// TIA Portal V19 export
DATA_BLOCK "Sim_SMOutputs_DB"   // DB9
// stored: InstanceOfName Sim_SMOutputs, InstanceOfType FB
"Sim_SMOutputs"
   // VAR
   //    VaccumPID { ExternalAccessible := 'False'; ExternalVisible := 'False'; ExternalWritable := 'False'} : "PidL";
   //    SteamPID { S7_SetPoint := 'True'} : "PidL";
   //    SimularDelay { S7_SetPoint := 'True'} : TON_TIME;
   //    FeedPID { S7_SetPoint := 'True'} : "PidL";
   //    LiSet : Bool := FALSE;
   //    LiSetM : Bool := FALSE;
   //    LevelInit : Real := 0.0;
   //    BrixInit : Real := 0.0;
   // END_VAR
BEGIN
   VaccumPID.AutModLi := TRUE;
   VaccumPID.ManModLi := FALSE;
   VaccumPID.LocModLi := FALSE;
   VaccumPID.OosModLi := FALSE;
   VaccumPID.ModLiOp := TRUE;
   VaccumPID.ResetLi := FALSE;
   VaccumPID.SPModLiOp := FALSE;
   VaccumPID.ExtModLi := FALSE;
   VaccumPID.IntModLi := FALSE;
   VaccumPID.PV := 950.0145;
   VaccumPID.PV_Norm.High := 2000.0;
   VaccumPID.PV_Norm.Low := 0.0;
   VaccumPID.MV_Norm.High := 100.0;
   VaccumPID.MV_Norm.Low := 0.0;
   VaccumPID.PV_Scale.High := 2000.0;
   VaccumPID.PV_Scale.Low := 0.0;
   VaccumPID.SPExt := 0.0;
   VaccumPID.SP_HiLim := 1000.0;
   VaccumPID.SP_LoLim := 0.0;
   VaccumPID.MV_HiLim := 100.0;
   VaccumPID.MV_LoLim := 0.0;
   VaccumPID.OosSafeMV := 0.0;
   VaccumPID.PV_unit := 1342;
   VaccumPID.MV_unit := 1342;
   VaccumPID.DataHMI.identName := '';
   VaccumPID.DataHMI.comment := '';
   VaccumPID.DataHMI.AutModOp := TRUE;
   VaccumPID.DataHMI.ManModOp := FALSE;
   VaccumPID.DataHMI.LocModOp := FALSE;
   VaccumPID.DataHMI.OosModOp := FALSE;
   VaccumPID.DataHMI.ResetOp := FALSE;
   VaccumPID.DataHMI.MonitorOn := FALSE;
   VaccumPID.DataHMI.ExtModOp := FALSE;
   VaccumPID.DataHMI.IntModOp := FALSE;
   VaccumPID.DataHMI.SpInt := 100.0;
   VaccumPID.DataHMI.Man := 0.0;
   VaccumPID.DataHMI.PermissionLog.AutModOpEn := FALSE;
   VaccumPID.DataHMI.PermissionLog.ManModOpEn := FALSE;
   VaccumPID.DataHMI.PermissionLog.LocModOpEn := FALSE;
   VaccumPID.DataHMI.PermissionLog.OosModOpEn := FALSE;
   VaccumPID.DataHMI.PermissionLog.ResetOpEn := TRUE;
   VaccumPID.DataHMI.PermissionLog.ExtModOpEn := FALSE;
   VaccumPID.DataHMI.PermissionLog.IntModOpEn := FALSE;
   VaccumPID.DataHMI.PermissionLog.Alarms.MsgSupEn := FALSE;
   VaccumPID.DataHMI.PermissionLog.Alarms.HiAlmSupEn := FALSE;
   VaccumPID.DataHMI.PermissionLog.Alarms.HiWrnSupEn := FALSE;
   VaccumPID.DataHMI.PermissionLog.Alarms.LoWrnSupEn := FALSE;
   VaccumPID.DataHMI.PermissionLog.Alarms.LoAlmSupEn := FALSE;
   VaccumPID.DataHMI.Status.OosAct := FALSE;
   VaccumPID.DataHMI.Status.LocAct := FALSE;
   VaccumPID.DataHMI.Status.ManAct := FALSE;
   VaccumPID.DataHMI.Status.AutAct := TRUE;
   VaccumPID.DataHMI.Status.SpExtAct := FALSE;
   VaccumPID.DataHMI.Status.Protection := FALSE;
   VaccumPID.DataHMI.Status.Intlock := TRUE;
   VaccumPID.DataHMI.Status.Permit := TRUE;
   VaccumPID.DataHMI.Status.TrackAct := TRUE;
   VaccumPID.DataHMI.Status.SP := 100.0;
   VaccumPID.DataHMI.Status.PV := 950.0145;
   VaccumPID.DataHMI.Status.ER := -845.0145;
   VaccumPID.DataHMI.Status.MV := 0.0;
   VaccumPID.DataHMI.Status.PVOpScale.High := 2000.0;
   VaccumPID.DataHMI.Status.PVOpScale.Low := 0.0;
   VaccumPID.DataHMI.Status.MVOpScale.High := 100.0;
   VaccumPID.DataHMI.Status.MVOpScale.Low := 0.0;
   VaccumPID.DataHMI.Status.SPIntLim.High := 0.0;
   VaccumPID.DataHMI.Status.SPIntLim.Low := 0.0;
   VaccumPID.DataHMI.Status.PV_unit := 1342;
   VaccumPID.DataHMI.Status.MV_unit := 1342;
   VaccumPID.DataHMI.PIDConfig.NegGain := TRUE;
   VaccumPID.DataHMI.PIDConfig.P_Sel := TRUE;
   VaccumPID.DataHMI.PIDConfig.I_Sel := TRUE;
   VaccumPID.DataHMI.PIDConfig.D_Sel := FALSE;
   VaccumPID.DataHMI.PIDConfig.Gain := -2.0;
   VaccumPID.DataHMI.PIDConfig.Ti := 80.0;
   VaccumPID.DataHMI.PIDConfig.Td := 0.0;
   VaccumPID.DataHMI.PIDConfig.DeadBW := 5.0;
   VaccumPID.DataHMI.Alarms.identName := '';
   VaccumPID.DataHMI.Alarms.comment := '';
   VaccumPID.DataHMI.Alarms.MsgSupOp := FALSE;
   VaccumPID.DataHMI.Alarms.PVScale.High := 2000.0;
   VaccumPID.DataHMI.Alarms.PVScale.Low := 0.0;
   VaccumPID.DataHMI.Alarms.HiAlmSupOp := FALSE;
   VaccumPID.DataHMI.Alarms.HiWrnSupOp := FALSE;
   VaccumPID.DataHMI.Alarms.LoWrnSupOp := FALSE;
   VaccumPID.DataHMI.Alarms.LoAlmSupOp := FALSE;
   VaccumPID.DataHMI.Alarms.PermissionLog.MsgSupEn := FALSE;
   VaccumPID.DataHMI.Alarms.PermissionLog.HiAlmSupEn := TRUE;
   VaccumPID.DataHMI.Alarms.PermissionLog.HiWrnSupEn := TRUE;
   VaccumPID.DataHMI.Alarms.PermissionLog.LoWrnSupEn := TRUE;
   VaccumPID.DataHMI.Alarms.PermissionLog.LoAlmSupEn := TRUE;
   VaccumPID.DataHMI.Alarms.Status.PV := 950.0145;
   VaccumPID.DataHMI.Alarms.Status.PV_unit := 1342;
   VaccumPID.DataHMI.Alarms.Status.PV_HiAlm := TRUE;
   VaccumPID.DataHMI.Alarms.Status.PV_HiWrn := TRUE;
   VaccumPID.DataHMI.Alarms.Status.PV_LoWrn := FALSE;
   VaccumPID.DataHMI.Alarms.Status.PV_LoAlm := FALSE;
   VaccumPID.DataHMI.Alarms.Status.MsgSup := FALSE;
   VaccumPID.Feature.Startup := TRUE;
   VaccumPID.Feature.MSSOff := TRUE;
   VaccumPID.Feature.FltOff := TRUE;
   VaccumPID.Feature.LocalMod := FALSE;
   VaccumPID.Permission.AutModOpEn := TRUE;
   VaccumPID.Permission.ManModOpEn := TRUE;
   VaccumPID.Permission.LocModOpEn := FALSE;
   VaccumPID.Permission.OosModOpEn := FALSE;
   VaccumPID.Permission.ResetOpEn := TRUE;
   VaccumPID.Permission.ExtModOpEn := FALSE;
   VaccumPID.Permission.IntModOpEn := TRUE;
   VaccumPID.Permission.Alarms.MsgSupEn := TRUE;
   VaccumPID.Permission.Alarms.HiAlmSupEn := TRUE;
   VaccumPID.Permission.Alarms.HiWrnSupEn := TRUE;
   VaccumPID.Permission.Alarms.LoWrnSupEn := TRUE;
   VaccumPID.Permission.Alarms.LoAlmSupEn := TRUE;
   VaccumPID.MSS := TRUE;
   VaccumPID.Trip := FALSE;
   VaccumPID.Permit := TRUE;
   VaccumPID.Intlock := TRUE;
   VaccumPID.Protect := TRUE;
   VaccumPID.TrackOn := TRUE;
   VaccumPID.Rbk := 0.0;
   VaccumPID.RbkHiTol := 3.0;
   VaccumPID.RbkLoTol := 3.0;
   VaccumPID.RbkMonTime := T#3S;
   VaccumPID.TrackVal := 0.0;
   VaccumPID.RunUpCyc := 3;
   VaccumPID.DisV := 0.0;
   VaccumPID.HiAlm := 95.0;
   VaccumPID.HiWrn := 90.0;
   VaccumPID.LoWrn := 10.0;
   VaccumPID.LoAlm := 5.0;
   VaccumPID.Hyst := 5.0;
   VaccumPID.AutAct := TRUE;
   VaccumPID.ManAct := FALSE;
   VaccumPID.LocAct := FALSE;
   VaccumPID.OosAct := FALSE;
   VaccumPID.MsgSup := TRUE;
   VaccumPID.AlarmError := FALSE;
   VaccumPID.MV := 0.0;
   VaccumPID.SPExtAct := FALSE;
   VaccumPID.SP := 100.0;
   VaccumPID.ER := -845.0145;
   VaccumPID.PVH_Alm := TRUE;
   VaccumPID.PVH_Wrn := TRUE;
   VaccumPID.PVL_Wrn := FALSE;
   VaccumPID.PVL_Alm := FALSE;
   VaccumPID.controller.COM_RST := FALSE;
   VaccumPID.controller.MAN_ON := TRUE;
   VaccumPID.controller.PVPER_ON := FALSE;
   VaccumPID.controller.P_SEL := TRUE;
   VaccumPID.controller.I_SEL := TRUE;
   VaccumPID.controller.INT_HOLD := FALSE;
   VaccumPID.controller.I_ITL_ON := FALSE;
   VaccumPID.controller.D_SEL := FALSE;
   VaccumPID.controller.CYCLE := T#200MS;
   VaccumPID.controller.SP_INT := 5.0;
   VaccumPID.controller.PV_IN := 47.50072;
   VaccumPID.controller.PV_PER := 16#0000;
   VaccumPID.controller.MAN := 0.0;
   VaccumPID.controller.GAIN := -2.0;
   VaccumPID.controller.TI := T#1M_20S;
   VaccumPID.controller.TD := T#10S;
   VaccumPID.controller.TM_LAG := T#2S;
   VaccumPID.controller.DEADB_W := 0.25;
   VaccumPID.controller.LMN_HLM := 100.0;
   VaccumPID.controller.LMN_LLM := 0.0;
   VaccumPID.controller.PV_FAC := 1.0;
   VaccumPID.controller.PV_OFF := 0.0;
   VaccumPID.controller.LMN_FAC := 1.0;
   VaccumPID.controller.LMN_OFF := 0.0;
   VaccumPID.controller.I_ITLVAL := 0.0;
   VaccumPID.controller.DISV := 0.0;
   VaccumPID.controller.LMN := 0.0;
   VaccumPID.controller.LMN_PER := 16#0000;
   VaccumPID.controller.QLMN_HLM := FALSE;
   VaccumPID.controller.QLMN_LLM := TRUE;
   VaccumPID.controller.LMN_P := 84.50145;
   VaccumPID.controller.LMN_I := -84.50145;
   VaccumPID.controller.LMN_D := 0.0;
   VaccumPID.controller.PV := 47.50072;
   VaccumPID.controller.ER := -42.25072;
   VaccumPID.controller.sInvAlt := 84.50145;
   VaccumPID.controller.sIanteilAlt := -84.50145;
   VaccumPID.controller.sRestInt := 0.0;
   VaccumPID.controller.sRestDif := 0.0;
   VaccumPID.controller.sRueck := 84.50145;
   VaccumPID.controller.sLmn := 0.0;
   VaccumPID.controller.sbArwHLmOn := FALSE;
   VaccumPID.controller.sbArwLLmOn := TRUE;
   VaccumPID.controller.sbILimOn := TRUE;
   VaccumPID.ModSelInt := 2;
   VaccumPID.stRestart := FALSE;
   VaccumPID.ResetLiLogic := FALSE;
   VaccumPID.ResetResult := FALSE;
   VaccumPID.stResetLiLogic := FALSE;
   VaccumPID.stMonErr := FALSE;
   VaccumPID.stTripErr := FALSE;
   VaccumPID.stProtErr := FALSE;
   VaccumPID.stMSS := FALSE;
   VaccumPID.stProt := FALSE;
   VaccumPID.stTrip := FALSE;
   VaccumPID.stLockFault := FALSE;
   VaccumPID.stRun := FALSE;
   VaccumPID.stExtMod := FALSE;
   VaccumPID.stAutoLogic := FALSE;
   VaccumPID.RuntimeMem := 16#0000_07DF_2C3D_9711;
   VaccumPID.RuntimeS := 0.200026255103497;
   VaccumPID.PVMon.Feature.Startup := TRUE;
   VaccumPID.PVMon.Enable := TRUE;
   VaccumPID.PVMon.Permission.MsgSupEn := TRUE;
   VaccumPID.PVMon.Permission.HiAlmSupEn := TRUE;
   VaccumPID.PVMon.Permission.HiWrnSupEn := TRUE;
   VaccumPID.PVMon.Permission.LoWrnSupEn := TRUE;
   VaccumPID.PVMon.Permission.LoAlmSupEn := TRUE;
   VaccumPID.PVMon.DataHMI.identName := '';
   VaccumPID.PVMon.DataHMI.comment := '';
   VaccumPID.PVMon.DataHMI.MsgSupOp := FALSE;
   VaccumPID.PVMon.DataHMI.PVScale.High := 2000.0;
   VaccumPID.PVMon.DataHMI.PVScale.Low := 0.0;
   VaccumPID.PVMon.DataHMI.HiAlmSupOp := FALSE;
   VaccumPID.PVMon.DataHMI.HiWrnSupOp := FALSE;
   VaccumPID.PVMon.DataHMI.LoWrnSupOp := FALSE;
   VaccumPID.PVMon.DataHMI.LoAlmSupOp := FALSE;
   VaccumPID.PVMon.DataHMI.PermissionLog.MsgSupEn := FALSE;
   VaccumPID.PVMon.DataHMI.PermissionLog.HiAlmSupEn := TRUE;
   VaccumPID.PVMon.DataHMI.PermissionLog.HiWrnSupEn := TRUE;
   VaccumPID.PVMon.DataHMI.PermissionLog.LoWrnSupEn := TRUE;
   VaccumPID.PVMon.DataHMI.PermissionLog.LoAlmSupEn := TRUE;
   VaccumPID.PVMon.DataHMI.Status.PV := 950.0145;
   VaccumPID.PVMon.DataHMI.Status.PV_unit := 1342;
   VaccumPID.PVMon.DataHMI.Status.PV_HiAlm := TRUE;
   VaccumPID.PVMon.DataHMI.Status.PV_HiWrn := TRUE;
   VaccumPID.PVMon.DataHMI.Status.PV_LoWrn := FALSE;
   VaccumPID.PVMon.DataHMI.Status.PV_LoAlm := FALSE;
   VaccumPID.PVMon.DataHMI.Status.MsgSup := FALSE;
   VaccumPID.PVMon.RunUpCyc := 3;
   VaccumPID.PVMon.PV := 950.0145;
   VaccumPID.PVMon.HiAlm := 95.0;
   VaccumPID.PVMon.HiWrn := 90.0;
   VaccumPID.PVMon.LoWrn := 10.0;
   VaccumPID.PVMon.LoAlm := 5.0;
   VaccumPID.PVMon.Hyst := 5.0;
   VaccumPID.PVMon.PV_unit := 1342;
   VaccumPID.PVMon.MsgErr := FALSE;
   VaccumPID.PVMon.MsgSup := FALSE;
   VaccumPID.PVMon.PVH_Alm := TRUE;
   VaccumPID.PVMon.PVH_Wrn := TRUE;
   VaccumPID.PVMon.PVL_Wrn := FALSE;
   VaccumPID.PVMon.PVL_Alm := FALSE;
   VaccumPID.PVMon.stRestart := FALSE;
   VaccumPID.PVMon.RunUpCounter := 0;
   VaccumPID.PVMon.pSIG1 := TRUE;
   VaccumPID.PVMon.pSIG2 := TRUE;
   VaccumPID.PVMon.pSIG3 := FALSE;
   VaccumPID.PVMon.pSIG4 := FALSE;
   VaccumPID.PVMon.pAlarm := TRUE;
   VaccumPID.RunUpCounter := 0;
   VaccumPID.pAlarm := TRUE;
   VaccumPID.stMSSErr := FALSE;
   VaccumPID.SPMod := FALSE;
   VaccumPID.SPSelInt := 0;
   VaccumPID.stErr := FALSE;
   VaccumPID.stDivErr := FALSE;
   VaccumPID.stNegGain := TRUE;
   VaccumPID.stGain := -2.0;
   VaccumPID.stTi := 0.0;
   VaccumPID.stTd := 0.0;
   VaccumPID.stPIDConfig.NegGain := TRUE;
   VaccumPID.stPIDConfig.P_Sel := TRUE;
   VaccumPID.stPIDConfig.I_Sel := TRUE;
   VaccumPID.stPIDConfig.D_Sel := FALSE;
   VaccumPID.stPIDConfig.Gain := -2.0;
   VaccumPID.stPIDConfig.Ti := 80.0;
   VaccumPID.stPIDConfig.Td := 0.0;
   VaccumPID.stPIDConfig.DeadBW := 5.0;
   VaccumPID.RbkMonitorTimer.PT := T#0MS;
   VaccumPID.RbkMonitorTimer.IN := FALSE;
   SteamPID.AutModLi := TRUE;
   SteamPID.ManModLi := FALSE;
   SteamPID.LocModLi := FALSE;
   SteamPID.OosModLi := FALSE;
   SteamPID.ModLiOp := TRUE;
   SteamPID.ResetLi := FALSE;
   SteamPID.SPModLiOp := TRUE;
   SteamPID.ExtModLi := TRUE;
   SteamPID.IntModLi := FALSE;
   SteamPID.PV := 0.0;
   SteamPID.PV_Norm.High := 100.0;
   SteamPID.PV_Norm.Low := 0.0;
   SteamPID.MV_Norm.High := 100.0;
   SteamPID.MV_Norm.Low := 0.0;
   SteamPID.PV_Scale.High := 100.0;
   SteamPID.PV_Scale.Low := 0.0;
   SteamPID.SPExt := 80.0;
   SteamPID.SP_HiLim := 100.0;
   SteamPID.SP_LoLim := 0.0;
   SteamPID.MV_HiLim := 100.0;
   SteamPID.MV_LoLim := 0.0;
   SteamPID.OosSafeMV := 0.0;
   SteamPID.PV_unit := 1342;
   SteamPID.MV_unit := 1342;
   SteamPID.DataHMI.identName := '';
   SteamPID.DataHMI.comment := '';
   SteamPID.DataHMI.AutModOp := TRUE;
   SteamPID.DataHMI.ManModOp := FALSE;
   SteamPID.DataHMI.LocModOp := FALSE;
   SteamPID.DataHMI.OosModOp := FALSE;
   SteamPID.DataHMI.ResetOp := FALSE;
   SteamPID.DataHMI.MonitorOn := FALSE;
   SteamPID.DataHMI.ExtModOp := FALSE;
   SteamPID.DataHMI.IntModOp := FALSE;
   SteamPID.DataHMI.SpInt := 80.0;
   SteamPID.DataHMI.Man := 0.0;
   SteamPID.DataHMI.PermissionLog.AutModOpEn := FALSE;
   SteamPID.DataHMI.PermissionLog.ManModOpEn := FALSE;
   SteamPID.DataHMI.PermissionLog.LocModOpEn := FALSE;
   SteamPID.DataHMI.PermissionLog.OosModOpEn := FALSE;
   SteamPID.DataHMI.PermissionLog.ResetOpEn := TRUE;
   SteamPID.DataHMI.PermissionLog.ExtModOpEn := FALSE;
   SteamPID.DataHMI.PermissionLog.IntModOpEn := FALSE;
   SteamPID.DataHMI.PermissionLog.Alarms.MsgSupEn := FALSE;
   SteamPID.DataHMI.PermissionLog.Alarms.HiAlmSupEn := FALSE;
   SteamPID.DataHMI.PermissionLog.Alarms.HiWrnSupEn := FALSE;
   SteamPID.DataHMI.PermissionLog.Alarms.LoWrnSupEn := FALSE;
   SteamPID.DataHMI.PermissionLog.Alarms.LoAlmSupEn := FALSE;
   SteamPID.DataHMI.Status.OosAct := FALSE;
   SteamPID.DataHMI.Status.LocAct := FALSE;
   SteamPID.DataHMI.Status.ManAct := FALSE;
   SteamPID.DataHMI.Status.AutAct := TRUE;
   SteamPID.DataHMI.Status.SpExtAct := TRUE;
   SteamPID.DataHMI.Status.Protection := FALSE;
   SteamPID.DataHMI.Status.Intlock := TRUE;
   SteamPID.DataHMI.Status.Permit := TRUE;
   SteamPID.DataHMI.Status.TrackAct := TRUE;
   SteamPID.DataHMI.Status.SP := 80.0;
   SteamPID.DataHMI.Status.PV := 0.0;
   SteamPID.DataHMI.Status.ER := 80.0;
   SteamPID.DataHMI.Status.MV := 0.0;
   SteamPID.DataHMI.Status.PVOpScale.High := 100.0;
   SteamPID.DataHMI.Status.PVOpScale.Low := 0.0;
   SteamPID.DataHMI.Status.MVOpScale.High := 100.0;
   SteamPID.DataHMI.Status.MVOpScale.Low := 0.0;
   SteamPID.DataHMI.Status.SPIntLim.High := 0.0;
   SteamPID.DataHMI.Status.SPIntLim.Low := 0.0;
   SteamPID.DataHMI.Status.PV_unit := 1342;
   SteamPID.DataHMI.Status.MV_unit := 1342;
   SteamPID.DataHMI.PIDConfig.NegGain := FALSE;
   SteamPID.DataHMI.PIDConfig.P_Sel := TRUE;
   SteamPID.DataHMI.PIDConfig.I_Sel := TRUE;
   SteamPID.DataHMI.PIDConfig.D_Sel := FALSE;
   SteamPID.DataHMI.PIDConfig.Gain := 2.0;
   SteamPID.DataHMI.PIDConfig.Ti := 80.0;
   SteamPID.DataHMI.PIDConfig.Td := 10.0;
   SteamPID.DataHMI.PIDConfig.DeadBW := 0.0;
   SteamPID.DataHMI.Alarms.identName := '';
   SteamPID.DataHMI.Alarms.comment := '';
   SteamPID.DataHMI.Alarms.MsgSupOp := FALSE;
   SteamPID.DataHMI.Alarms.PVScale.High := 100.0;
   SteamPID.DataHMI.Alarms.PVScale.Low := 0.0;
   SteamPID.DataHMI.Alarms.HiAlmSupOp := FALSE;
   SteamPID.DataHMI.Alarms.HiWrnSupOp := FALSE;
   SteamPID.DataHMI.Alarms.LoWrnSupOp := FALSE;
   SteamPID.DataHMI.Alarms.LoAlmSupOp := FALSE;
   SteamPID.DataHMI.Alarms.PermissionLog.MsgSupEn := FALSE;
   SteamPID.DataHMI.Alarms.PermissionLog.HiAlmSupEn := TRUE;
   SteamPID.DataHMI.Alarms.PermissionLog.HiWrnSupEn := TRUE;
   SteamPID.DataHMI.Alarms.PermissionLog.LoWrnSupEn := TRUE;
   SteamPID.DataHMI.Alarms.PermissionLog.LoAlmSupEn := TRUE;
   SteamPID.DataHMI.Alarms.Status.PV := 0.0;
   SteamPID.DataHMI.Alarms.Status.PV_unit := 1342;
   SteamPID.DataHMI.Alarms.Status.PV_HiAlm := FALSE;
   SteamPID.DataHMI.Alarms.Status.PV_HiWrn := FALSE;
   SteamPID.DataHMI.Alarms.Status.PV_LoWrn := TRUE;
   SteamPID.DataHMI.Alarms.Status.PV_LoAlm := TRUE;
   SteamPID.DataHMI.Alarms.Status.MsgSup := FALSE;
   SteamPID.Feature.Startup := TRUE;
   SteamPID.Feature.MSSOff := TRUE;
   SteamPID.Feature.FltOff := TRUE;
   SteamPID.Feature.LocalMod := FALSE;
   SteamPID.Permission.AutModOpEn := TRUE;
   SteamPID.Permission.ManModOpEn := TRUE;
   SteamPID.Permission.LocModOpEn := FALSE;
   SteamPID.Permission.OosModOpEn := FALSE;
   SteamPID.Permission.ResetOpEn := TRUE;
   SteamPID.Permission.ExtModOpEn := FALSE;
   SteamPID.Permission.IntModOpEn := TRUE;
   SteamPID.Permission.Alarms.MsgSupEn := TRUE;
   SteamPID.Permission.Alarms.HiAlmSupEn := TRUE;
   SteamPID.Permission.Alarms.HiWrnSupEn := TRUE;
   SteamPID.Permission.Alarms.LoWrnSupEn := TRUE;
   SteamPID.Permission.Alarms.LoAlmSupEn := TRUE;
   SteamPID.MSS := TRUE;
   SteamPID.Trip := FALSE;
   SteamPID.Permit := TRUE;
   SteamPID.Intlock := TRUE;
   SteamPID.Protect := TRUE;
   SteamPID.TrackOn := TRUE;
   SteamPID.Rbk := 0.0;
   SteamPID.RbkHiTol := 3.0;
   SteamPID.RbkLoTol := 3.0;
   SteamPID.RbkMonTime := T#3S;
   SteamPID.TrackVal := 0.0;
   SteamPID.RunUpCyc := 3;
   SteamPID.DisV := 0.0;
   SteamPID.HiAlm := 95.0;
   SteamPID.HiWrn := 90.0;
   SteamPID.LoWrn := 10.0;
   SteamPID.LoAlm := 5.0;
   SteamPID.Hyst := 5.0;
   SteamPID.AutAct := TRUE;
   SteamPID.ManAct := FALSE;
   SteamPID.LocAct := FALSE;
   SteamPID.OosAct := FALSE;
   SteamPID.MsgSup := TRUE;
   SteamPID.AlarmError := FALSE;
   SteamPID.MV := 0.0;
   SteamPID.SPExtAct := TRUE;
   SteamPID.SP := 80.0;
   SteamPID.ER := 80.0;
   SteamPID.PVH_Alm := FALSE;
   SteamPID.PVH_Wrn := FALSE;
   SteamPID.PVL_Wrn := TRUE;
   SteamPID.PVL_Alm := TRUE;
   SteamPID.controller.COM_RST := FALSE;
   SteamPID.controller.MAN_ON := TRUE;
   SteamPID.controller.PVPER_ON := FALSE;
   SteamPID.controller.P_SEL := TRUE;
   SteamPID.controller.I_SEL := TRUE;
   SteamPID.controller.INT_HOLD := FALSE;
   SteamPID.controller.I_ITL_ON := FALSE;
   SteamPID.controller.D_SEL := FALSE;
   SteamPID.controller.CYCLE := T#200MS;
   SteamPID.controller.SP_INT := 80.0;
   SteamPID.controller.PV_IN := 0.0;
   SteamPID.controller.PV_PER := 16#0000;
   SteamPID.controller.MAN := 0.0;
   SteamPID.controller.GAIN := 2.0;
   SteamPID.controller.TI := T#1M_20S;
   SteamPID.controller.TD := T#10S;
   SteamPID.controller.TM_LAG := T#2S;
   SteamPID.controller.DEADB_W := 0.0;
   SteamPID.controller.LMN_HLM := 100.0;
   SteamPID.controller.LMN_LLM := 0.0;
   SteamPID.controller.PV_FAC := 1.0;
   SteamPID.controller.PV_OFF := 0.0;
   SteamPID.controller.LMN_FAC := 1.0;
   SteamPID.controller.LMN_OFF := 0.0;
   SteamPID.controller.I_ITLVAL := 0.0;
   SteamPID.controller.DISV := 0.0;
   SteamPID.controller.LMN := 0.0;
   SteamPID.controller.LMN_PER := 16#0000;
   SteamPID.controller.QLMN_HLM := FALSE;
   SteamPID.controller.QLMN_LLM := TRUE;
   SteamPID.controller.LMN_P := 160.0;
   SteamPID.controller.LMN_I := -160.0;
   SteamPID.controller.LMN_D := 0.0;
   SteamPID.controller.PV := 0.0;
   SteamPID.controller.ER := 80.0;
   SteamPID.controller.sInvAlt := 160.0;
   SteamPID.controller.sIanteilAlt := -160.0;
   SteamPID.controller.sRestInt := 0.0;
   SteamPID.controller.sRestDif := 0.0;
   SteamPID.controller.sRueck := 160.0;
   SteamPID.controller.sLmn := 0.0;
   SteamPID.controller.sbArwHLmOn := FALSE;
   SteamPID.controller.sbArwLLmOn := TRUE;
   SteamPID.controller.sbILimOn := TRUE;
   SteamPID.ModSelInt := 2;
   SteamPID.stRestart := FALSE;
   SteamPID.ResetLiLogic := FALSE;
   SteamPID.ResetResult := FALSE;
   SteamPID.stResetLiLogic := FALSE;
   SteamPID.stMonErr := FALSE;
   SteamPID.stTripErr := FALSE;
   SteamPID.stProtErr := FALSE;
   SteamPID.stMSS := FALSE;
   SteamPID.stProt := FALSE;
   SteamPID.stTrip := FALSE;
   SteamPID.stLockFault := FALSE;
   SteamPID.stRun := FALSE;
   SteamPID.stExtMod := FALSE;
   SteamPID.stAutoLogic := FALSE;
   SteamPID.RuntimeMem := 16#0000_07DF_2C3F_7F80;
   SteamPID.RuntimeS := 0.200023537350218;
   SteamPID.PVMon.Feature.Startup := TRUE;
   SteamPID.PVMon.Enable := TRUE;
   SteamPID.PVMon.Permission.MsgSupEn := TRUE;
   SteamPID.PVMon.Permission.HiAlmSupEn := TRUE;
   SteamPID.PVMon.Permission.HiWrnSupEn := TRUE;
   SteamPID.PVMon.Permission.LoWrnSupEn := TRUE;
   SteamPID.PVMon.Permission.LoAlmSupEn := TRUE;
   SteamPID.PVMon.DataHMI.identName := '';
   SteamPID.PVMon.DataHMI.comment := '';
   SteamPID.PVMon.DataHMI.MsgSupOp := FALSE;
   SteamPID.PVMon.DataHMI.PVScale.High := 100.0;
   SteamPID.PVMon.DataHMI.PVScale.Low := 0.0;
   SteamPID.PVMon.DataHMI.HiAlmSupOp := FALSE;
   SteamPID.PVMon.DataHMI.HiWrnSupOp := FALSE;
   SteamPID.PVMon.DataHMI.LoWrnSupOp := FALSE;
   SteamPID.PVMon.DataHMI.LoAlmSupOp := FALSE;
   SteamPID.PVMon.DataHMI.PermissionLog.MsgSupEn := FALSE;
   SteamPID.PVMon.DataHMI.PermissionLog.HiAlmSupEn := TRUE;
   SteamPID.PVMon.DataHMI.PermissionLog.HiWrnSupEn := TRUE;
   SteamPID.PVMon.DataHMI.PermissionLog.LoWrnSupEn := TRUE;
   SteamPID.PVMon.DataHMI.PermissionLog.LoAlmSupEn := TRUE;
   SteamPID.PVMon.DataHMI.Status.PV := 0.0;
   SteamPID.PVMon.DataHMI.Status.PV_unit := 1342;
   SteamPID.PVMon.DataHMI.Status.PV_HiAlm := FALSE;
   SteamPID.PVMon.DataHMI.Status.PV_HiWrn := FALSE;
   SteamPID.PVMon.DataHMI.Status.PV_LoWrn := TRUE;
   SteamPID.PVMon.DataHMI.Status.PV_LoAlm := TRUE;
   SteamPID.PVMon.DataHMI.Status.MsgSup := FALSE;
   SteamPID.PVMon.RunUpCyc := 3;
   SteamPID.PVMon.PV := 0.0;
   SteamPID.PVMon.HiAlm := 95.0;
   SteamPID.PVMon.HiWrn := 90.0;
   SteamPID.PVMon.LoWrn := 10.0;
   SteamPID.PVMon.LoAlm := 5.0;
   SteamPID.PVMon.Hyst := 5.0;
   SteamPID.PVMon.PV_unit := 1342;
   SteamPID.PVMon.MsgErr := FALSE;
   SteamPID.PVMon.MsgSup := FALSE;
   SteamPID.PVMon.PVH_Alm := FALSE;
   SteamPID.PVMon.PVH_Wrn := FALSE;
   SteamPID.PVMon.PVL_Wrn := TRUE;
   SteamPID.PVMon.PVL_Alm := TRUE;
   SteamPID.PVMon.stRestart := FALSE;
   SteamPID.PVMon.RunUpCounter := 0;
   SteamPID.PVMon.pSIG1 := FALSE;
   SteamPID.PVMon.pSIG2 := FALSE;
   SteamPID.PVMon.pSIG3 := TRUE;
   SteamPID.PVMon.pSIG4 := TRUE;
   SteamPID.PVMon.pAlarm := TRUE;
   SteamPID.RunUpCounter := 0;
   SteamPID.pAlarm := TRUE;
   SteamPID.stMSSErr := FALSE;
   SteamPID.SPMod := FALSE;
   SteamPID.SPSelInt := 2;
   SteamPID.stErr := FALSE;
   SteamPID.stDivErr := FALSE;
   SteamPID.stNegGain := FALSE;
   SteamPID.stGain := 2.0;
   SteamPID.stTi := 0.0;
   SteamPID.stTd := 0.0;
   SteamPID.stPIDConfig.NegGain := FALSE;
   SteamPID.stPIDConfig.P_Sel := TRUE;
   SteamPID.stPIDConfig.I_Sel := TRUE;
   SteamPID.stPIDConfig.D_Sel := FALSE;
   SteamPID.stPIDConfig.Gain := 2.0;
   SteamPID.stPIDConfig.Ti := 80.0;
   SteamPID.stPIDConfig.Td := 10.0;
   SteamPID.stPIDConfig.DeadBW := 0.0;
   SteamPID.RbkMonitorTimer.PT := T#0MS;
   SteamPID.RbkMonitorTimer.IN := FALSE;
   SimularDelay.PT := T#2S;
   SimularDelay.IN := TRUE;
   FeedPID.AutModLi := TRUE;
   FeedPID.ManModLi := FALSE;
   FeedPID.LocModLi := FALSE;
   FeedPID.OosModLi := FALSE;
   FeedPID.ModLiOp := TRUE;
   FeedPID.ResetLi := FALSE;
   FeedPID.SPModLiOp := FALSE;
   FeedPID.ExtModLi := FALSE;
   FeedPID.IntModLi := FALSE;
   FeedPID.PV := 0.0;
   FeedPID.PV_Norm.High := 100.0;
   FeedPID.PV_Norm.Low := 0.0;
   FeedPID.MV_Norm.High := 100.0;
   FeedPID.MV_Norm.Low := 0.0;
   FeedPID.PV_Scale.High := 100.0;
   FeedPID.PV_Scale.Low := 0.0;
   FeedPID.SPExt := 0.0;
   FeedPID.SP_HiLim := 100.0;
   FeedPID.SP_LoLim := 0.0;
   FeedPID.MV_HiLim := 100.0;
   FeedPID.MV_LoLim := 0.0;
   FeedPID.OosSafeMV := 0.0;
   FeedPID.PV_unit := 1342;
   FeedPID.MV_unit := 1342;
   FeedPID.DataHMI.identName := '';
   FeedPID.DataHMI.comment := '';
   FeedPID.DataHMI.AutModOp := TRUE;
   FeedPID.DataHMI.ManModOp := FALSE;
   FeedPID.DataHMI.LocModOp := FALSE;
   FeedPID.DataHMI.OosModOp := FALSE;
   FeedPID.DataHMI.ResetOp := FALSE;
   FeedPID.DataHMI.MonitorOn := FALSE;
   FeedPID.DataHMI.ExtModOp := FALSE;
   FeedPID.DataHMI.IntModOp := FALSE;
   FeedPID.DataHMI.SpInt := 85.2033;
   FeedPID.DataHMI.Man := 0.0;
   FeedPID.DataHMI.PermissionLog.AutModOpEn := FALSE;
   FeedPID.DataHMI.PermissionLog.ManModOpEn := FALSE;
   FeedPID.DataHMI.PermissionLog.LocModOpEn := FALSE;
   FeedPID.DataHMI.PermissionLog.OosModOpEn := FALSE;
   FeedPID.DataHMI.PermissionLog.ResetOpEn := TRUE;
   FeedPID.DataHMI.PermissionLog.ExtModOpEn := FALSE;
   FeedPID.DataHMI.PermissionLog.IntModOpEn := FALSE;
   FeedPID.DataHMI.PermissionLog.Alarms.MsgSupEn := FALSE;
   FeedPID.DataHMI.PermissionLog.Alarms.HiAlmSupEn := FALSE;
   FeedPID.DataHMI.PermissionLog.Alarms.HiWrnSupEn := FALSE;
   FeedPID.DataHMI.PermissionLog.Alarms.LoWrnSupEn := FALSE;
   FeedPID.DataHMI.PermissionLog.Alarms.LoAlmSupEn := FALSE;
   FeedPID.DataHMI.Status.OosAct := FALSE;
   FeedPID.DataHMI.Status.LocAct := FALSE;
   FeedPID.DataHMI.Status.ManAct := FALSE;
   FeedPID.DataHMI.Status.AutAct := TRUE;
   FeedPID.DataHMI.Status.SpExtAct := FALSE;
   FeedPID.DataHMI.Status.Protection := FALSE;
   FeedPID.DataHMI.Status.Intlock := TRUE;
   FeedPID.DataHMI.Status.Permit := TRUE;
   FeedPID.DataHMI.Status.TrackAct := TRUE;
   FeedPID.DataHMI.Status.SP := 85.2033;
   FeedPID.DataHMI.Status.PV := 0.0;
   FeedPID.DataHMI.Status.ER := 85.2033;
   FeedPID.DataHMI.Status.MV := 0.0;
   FeedPID.DataHMI.Status.PVOpScale.High := 100.0;
   FeedPID.DataHMI.Status.PVOpScale.Low := 0.0;
   FeedPID.DataHMI.Status.MVOpScale.High := 100.0;
   FeedPID.DataHMI.Status.MVOpScale.Low := 0.0;
   FeedPID.DataHMI.Status.SPIntLim.High := 0.0;
   FeedPID.DataHMI.Status.SPIntLim.Low := 0.0;
   FeedPID.DataHMI.Status.PV_unit := 1342;
   FeedPID.DataHMI.Status.MV_unit := 1342;
   FeedPID.DataHMI.PIDConfig.NegGain := FALSE;
   FeedPID.DataHMI.PIDConfig.P_Sel := TRUE;
   FeedPID.DataHMI.PIDConfig.I_Sel := TRUE;
   FeedPID.DataHMI.PIDConfig.D_Sel := FALSE;
   FeedPID.DataHMI.PIDConfig.Gain := 2.0;
   FeedPID.DataHMI.PIDConfig.Ti := 20.0;
   FeedPID.DataHMI.PIDConfig.Td := 10.0;
   FeedPID.DataHMI.PIDConfig.DeadBW := 0.0;
   FeedPID.DataHMI.Alarms.identName := '';
   FeedPID.DataHMI.Alarms.comment := '';
   FeedPID.DataHMI.Alarms.MsgSupOp := FALSE;
   FeedPID.DataHMI.Alarms.PVScale.High := 100.0;
   FeedPID.DataHMI.Alarms.PVScale.Low := 0.0;
   FeedPID.DataHMI.Alarms.HiAlmSupOp := FALSE;
   FeedPID.DataHMI.Alarms.HiWrnSupOp := FALSE;
   FeedPID.DataHMI.Alarms.LoWrnSupOp := FALSE;
   FeedPID.DataHMI.Alarms.LoAlmSupOp := FALSE;
   FeedPID.DataHMI.Alarms.PermissionLog.MsgSupEn := FALSE;
   FeedPID.DataHMI.Alarms.PermissionLog.HiAlmSupEn := TRUE;
   FeedPID.DataHMI.Alarms.PermissionLog.HiWrnSupEn := TRUE;
   FeedPID.DataHMI.Alarms.PermissionLog.LoWrnSupEn := TRUE;
   FeedPID.DataHMI.Alarms.PermissionLog.LoAlmSupEn := TRUE;
   FeedPID.DataHMI.Alarms.Status.PV := 0.0;
   FeedPID.DataHMI.Alarms.Status.PV_unit := 1342;
   FeedPID.DataHMI.Alarms.Status.PV_HiAlm := FALSE;
   FeedPID.DataHMI.Alarms.Status.PV_HiWrn := FALSE;
   FeedPID.DataHMI.Alarms.Status.PV_LoWrn := TRUE;
   FeedPID.DataHMI.Alarms.Status.PV_LoAlm := TRUE;
   FeedPID.DataHMI.Alarms.Status.MsgSup := FALSE;
   FeedPID.Feature.Startup := TRUE;
   FeedPID.Feature.MSSOff := TRUE;
   FeedPID.Feature.FltOff := TRUE;
   FeedPID.Feature.LocalMod := FALSE;
   FeedPID.Permission.AutModOpEn := TRUE;
   FeedPID.Permission.ManModOpEn := TRUE;
   FeedPID.Permission.LocModOpEn := FALSE;
   FeedPID.Permission.OosModOpEn := FALSE;
   FeedPID.Permission.ResetOpEn := TRUE;
   FeedPID.Permission.ExtModOpEn := FALSE;
   FeedPID.Permission.IntModOpEn := TRUE;
   FeedPID.Permission.Alarms.MsgSupEn := TRUE;
   FeedPID.Permission.Alarms.HiAlmSupEn := TRUE;
   FeedPID.Permission.Alarms.HiWrnSupEn := TRUE;
   FeedPID.Permission.Alarms.LoWrnSupEn := TRUE;
   FeedPID.Permission.Alarms.LoAlmSupEn := TRUE;
   FeedPID.MSS := TRUE;
   FeedPID.Trip := FALSE;
   FeedPID.Permit := TRUE;
   FeedPID.Intlock := TRUE;
   FeedPID.Protect := TRUE;
   FeedPID.TrackOn := TRUE;
   FeedPID.Rbk := 0.0;
   FeedPID.RbkHiTol := 3.0;
   FeedPID.RbkLoTol := 3.0;
   FeedPID.RbkMonTime := T#3S;
   FeedPID.TrackVal := 0.0;
   FeedPID.RunUpCyc := 3;
   FeedPID.DisV := 0.0;
   FeedPID.HiAlm := 95.0;
   FeedPID.HiWrn := 90.0;
   FeedPID.LoWrn := 10.0;
   FeedPID.LoAlm := 5.0;
   FeedPID.Hyst := 5.0;
   FeedPID.AutAct := TRUE;
   FeedPID.ManAct := FALSE;
   FeedPID.LocAct := FALSE;
   FeedPID.OosAct := FALSE;
   FeedPID.MsgSup := TRUE;
   FeedPID.AlarmError := FALSE;
   FeedPID.MV := 0.0;
   FeedPID.SPExtAct := FALSE;
   FeedPID.SP := 85.2033;
   FeedPID.ER := 85.2033;
   FeedPID.PVH_Alm := FALSE;
   FeedPID.PVH_Wrn := FALSE;
   FeedPID.PVL_Wrn := TRUE;
   FeedPID.PVL_Alm := TRUE;
   FeedPID.controller.COM_RST := FALSE;
   FeedPID.controller.MAN_ON := TRUE;
   FeedPID.controller.PVPER_ON := FALSE;
   FeedPID.controller.P_SEL := TRUE;
   FeedPID.controller.I_SEL := TRUE;
   FeedPID.controller.INT_HOLD := FALSE;
   FeedPID.controller.I_ITL_ON := FALSE;
   FeedPID.controller.D_SEL := FALSE;
   FeedPID.controller.CYCLE := T#200MS;
   FeedPID.controller.SP_INT := 85.2033;
   FeedPID.controller.PV_IN := 0.0;
   FeedPID.controller.PV_PER := 16#0000;
   FeedPID.controller.MAN := 0.0;
   FeedPID.controller.GAIN := 2.0;
   FeedPID.controller.TI := T#20S;
   FeedPID.controller.TD := T#10S;
   FeedPID.controller.TM_LAG := T#2S;
   FeedPID.controller.DEADB_W := 0.0;
   FeedPID.controller.LMN_HLM := 100.0;
   FeedPID.controller.LMN_LLM := 0.0;
   FeedPID.controller.PV_FAC := 1.0;
   FeedPID.controller.PV_OFF := 0.0;
   FeedPID.controller.LMN_FAC := 1.0;
   FeedPID.controller.LMN_OFF := 0.0;
   FeedPID.controller.I_ITLVAL := 0.0;
   FeedPID.controller.DISV := 0.0;
   FeedPID.controller.LMN := 0.0;
   FeedPID.controller.LMN_PER := 16#0000;
   FeedPID.controller.QLMN_HLM := FALSE;
   FeedPID.controller.QLMN_LLM := TRUE;
   FeedPID.controller.LMN_P := 170.4066;
   FeedPID.controller.LMN_I := -170.4066;
   FeedPID.controller.LMN_D := 0.0;
   FeedPID.controller.PV := 0.0;
   FeedPID.controller.ER := 85.2033;
   FeedPID.controller.sInvAlt := 170.4066;
   FeedPID.controller.sIanteilAlt := -170.4066;
   FeedPID.controller.sRestInt := 0.0;
   FeedPID.controller.sRestDif := 0.0;
   FeedPID.controller.sRueck := 170.4066;
   FeedPID.controller.sLmn := 0.0;
   FeedPID.controller.sbArwHLmOn := FALSE;
   FeedPID.controller.sbArwLLmOn := TRUE;
   FeedPID.controller.sbILimOn := TRUE;
   FeedPID.ModSelInt := 2;
   FeedPID.stRestart := FALSE;
   FeedPID.ResetLiLogic := FALSE;
   FeedPID.ResetResult := FALSE;
   FeedPID.stResetLiLogic := FALSE;
   FeedPID.stMonErr := FALSE;
   FeedPID.stTripErr := FALSE;
   FeedPID.stProtErr := FALSE;
   FeedPID.stMSS := FALSE;
   FeedPID.stProt := FALSE;
   FeedPID.stTrip := FALSE;
   FeedPID.stLockFault := FALSE;
   FeedPID.stRun := FALSE;
   FeedPID.stExtMod := FALSE;
   FeedPID.stAutoLogic := FALSE;
   FeedPID.RuntimeMem := 16#0000_07DF_2C40_BF76;
   FeedPID.RuntimeS := 0.200024909247694;
   FeedPID.PVMon.Feature.Startup := TRUE;
   FeedPID.PVMon.Enable := TRUE;
   FeedPID.PVMon.Permission.MsgSupEn := TRUE;
   FeedPID.PVMon.Permission.HiAlmSupEn := TRUE;
   FeedPID.PVMon.Permission.HiWrnSupEn := TRUE;
   FeedPID.PVMon.Permission.LoWrnSupEn := TRUE;
   FeedPID.PVMon.Permission.LoAlmSupEn := TRUE;
   FeedPID.PVMon.DataHMI.identName := '';
   FeedPID.PVMon.DataHMI.comment := '';
   FeedPID.PVMon.DataHMI.MsgSupOp := FALSE;
   FeedPID.PVMon.DataHMI.PVScale.High := 100.0;
   FeedPID.PVMon.DataHMI.PVScale.Low := 0.0;
   FeedPID.PVMon.DataHMI.HiAlmSupOp := FALSE;
   FeedPID.PVMon.DataHMI.HiWrnSupOp := FALSE;
   FeedPID.PVMon.DataHMI.LoWrnSupOp := FALSE;
   FeedPID.PVMon.DataHMI.LoAlmSupOp := FALSE;
   FeedPID.PVMon.DataHMI.PermissionLog.MsgSupEn := FALSE;
   FeedPID.PVMon.DataHMI.PermissionLog.HiAlmSupEn := TRUE;
   FeedPID.PVMon.DataHMI.PermissionLog.HiWrnSupEn := TRUE;
   FeedPID.PVMon.DataHMI.PermissionLog.LoWrnSupEn := TRUE;
   FeedPID.PVMon.DataHMI.PermissionLog.LoAlmSupEn := TRUE;
   FeedPID.PVMon.DataHMI.Status.PV := 0.0;
   FeedPID.PVMon.DataHMI.Status.PV_unit := 1342;
   FeedPID.PVMon.DataHMI.Status.PV_HiAlm := FALSE;
   FeedPID.PVMon.DataHMI.Status.PV_HiWrn := FALSE;
   FeedPID.PVMon.DataHMI.Status.PV_LoWrn := TRUE;
   FeedPID.PVMon.DataHMI.Status.PV_LoAlm := TRUE;
   FeedPID.PVMon.DataHMI.Status.MsgSup := FALSE;
   FeedPID.PVMon.RunUpCyc := 3;
   FeedPID.PVMon.PV := 0.0;
   FeedPID.PVMon.HiAlm := 95.0;
   FeedPID.PVMon.HiWrn := 90.0;
   FeedPID.PVMon.LoWrn := 10.0;
   FeedPID.PVMon.LoAlm := 5.0;
   FeedPID.PVMon.Hyst := 5.0;
   FeedPID.PVMon.PV_unit := 1342;
   FeedPID.PVMon.MsgErr := FALSE;
   FeedPID.PVMon.MsgSup := FALSE;
   FeedPID.PVMon.PVH_Alm := FALSE;
   FeedPID.PVMon.PVH_Wrn := FALSE;
   FeedPID.PVMon.PVL_Wrn := TRUE;
   FeedPID.PVMon.PVL_Alm := TRUE;
   FeedPID.PVMon.stRestart := FALSE;
   FeedPID.PVMon.RunUpCounter := 0;
   FeedPID.PVMon.pSIG1 := FALSE;
   FeedPID.PVMon.pSIG2 := FALSE;
   FeedPID.PVMon.pSIG3 := TRUE;
   FeedPID.PVMon.pSIG4 := TRUE;
   FeedPID.PVMon.pAlarm := TRUE;
   FeedPID.RunUpCounter := 0;
   FeedPID.pAlarm := TRUE;
   FeedPID.stMSSErr := FALSE;
   FeedPID.SPMod := FALSE;
   FeedPID.SPSelInt := 0;
   FeedPID.stErr := FALSE;
   FeedPID.stDivErr := FALSE;
   FeedPID.stNegGain := FALSE;
   FeedPID.stGain := 2.0;
   FeedPID.stTi := 0.0;
   FeedPID.stTd := 0.0;
   FeedPID.stPIDConfig.NegGain := FALSE;
   FeedPID.stPIDConfig.P_Sel := TRUE;
   FeedPID.stPIDConfig.I_Sel := TRUE;
   FeedPID.stPIDConfig.D_Sel := FALSE;
   FeedPID.stPIDConfig.Gain := 2.0;
   FeedPID.stPIDConfig.Ti := 20.0;
   FeedPID.stPIDConfig.Td := 10.0;
   FeedPID.stPIDConfig.DeadBW := 0.0;
   FeedPID.RbkMonitorTimer.PT := T#0MS;
   FeedPID.RbkMonitorTimer.IN := FALSE;
END_DATA_BLOCK
